Fanuc KAREL source: KO00018.KL

PROGRAM KO00018
%NOLOCKGROUP
VAR
  P1: XYZWPREXT
  P2: XYZWPREXT
  P3: XYZWPREXT
  OUT: XYZWPR
BEGIN
  OUT = FRAME(P1, P2, P3)
END KO00018
